(* IEC 61131-3 sources: Lasal-MCP/examples/SampleSource/5_ClassInputOutputSolution/Stations/MachineControl/MachineControl/Class/ValuesForComponents, 1 file *)

(* ---- ValuesForComponents.st ---- *)
(*!
<Class
	Name               = "ValuesForComponents"
	Revision           = "0.0"
	RealtimeTask       = "false"
	CyclicTask         = "false"
	BackgroundTask     = "false"
	Sigmatek           = "false"
	OSInterface        = "false"
	HighPriority       = "false"
	Automatic          = "false"
	UpdateMode         = "Prescan"
	SharedCommandTable = "true"
	Objectsize         = "(514,120)">
	<Channels>
		<Server Name="MyBar" Visualized="true" Initialize="false" WriteProtected="false" Retentive="false"/>
		<Server Name="MyDate" Visualized="true" Initialize="false" WriteProtected="false" Retentive="false"/>
		<Server Name="MyEnumeration" Visualized="true" Initialize="false" WriteProtected="false" Retentive="false"/>
		<Server Name="MyIPAddress" Visualized="true" Initialize="false" WriteProtected="false" Retentive="false"/>
		<Server Name="MyMenu" Visualized="true" Initialize="false" WriteProtected="false" Retentive="false"/>
		<Server Name="MyTime" Visualized="true" Initialize="false" WriteProtected="false" Retentive="false"/>
	</Channels>
</Class>
*)
ValuesForComponents : CLASS
	TYPE
	  t_MACHINE_STEPS :  //! <Type Public="true" Name="t_MACHINE_STEPS"/>
	  (
	    _Machine_Steps_NOOP,
	    _Machine_Steps_IDLE,
	    _Machine_Steps_HAND,
	    _Machine_Steps_AUTO
	  )$UDINT;
	END_TYPE
  //Servers:
	MyTime 	: SvrChCmd_DINT;
	MyDate 	: SvrCh_DINT;
	MyIPAddress 	: SvrCh_HDINT;
	MyEnumeration 	: SvrCh_t_MACHINE_STEPS_PTofCls_ValuesForComponents;
	MyMenu 	: SvrCh_DINT;
	MyBar 	: SvrCh_DINT;
  //Clients:
  //Variables:
  //Functions:
  //Tables:
	FUNCTION @STD
		VAR_OUTPUT
			ret_code	: CONFSTATES;
		END_VAR;
	FUNCTION GLOBAL TAB @CT_;
END_CLASS;
